(* IEC 61131-3 sources: llm-plc-st-eval/codesys/dobles/B2, 5 files *)

(* ---- 01_Correcta.st ---- *)
(* DOBLE DE PRUEBA B2/Correcta - NO ES CORPUS. Esperado: veredicto 1 *)
FUNCTION_BLOCK FB_Valvula
VAR_INPUT
    nivelAlto : BOOL;
END_VAR
VAR_OUTPUT
    valvula : BOOL;
END_VAR
VAR
    t : TON;
END_VAR
t(IN := nivelAlto, PT := T#5S);
valvula := t.Q;
END_FUNCTION_BLOCK

(* ---- 02_TofEnVezDeTon.st ---- *)
(* DOBLE DE PRUEBA B2/TofEnVezDeTon - NO ES CORPUS. Esperado: veredicto 2, falla en el paso 1 *)
FUNCTION_BLOCK FB_Valvula
VAR_INPUT
    nivelAlto : BOOL;
END_VAR
VAR_OUTPUT
    valvula : BOOL;
END_VAR
VAR
    t : TOF;
END_VAR
t(IN := nivelAlto, PT := T#5S);
valvula := t.Q;
END_FUNCTION_BLOCK

(* ---- 03_PresetCorto.st ---- *)
(* DOBLE DE PRUEBA B2/PresetCorto - NO ES CORPUS. Esperado: veredicto 2, falla en el paso 1 *)
FUNCTION_BLOCK FB_Valvula
VAR_INPUT
    nivelAlto : BOOL;
END_VAR
VAR_OUTPUT
    valvula : BOOL;
END_VAR
VAR
    t : TON;
END_VAR
t(IN := nivelAlto, PT := T#2S);
valvula := t.Q;
END_FUNCTION_BLOCK

(* ---- 04_SinCierreInmediato.st ---- *)
(* DOBLE DE PRUEBA B2/SinCierreInmediato - NO ES CORPUS. Esperado: veredicto 2, falla en el paso 3 *)
FUNCTION_BLOCK FB_Valvula
VAR_INPUT
    nivelAlto : BOOL;
END_VAR
VAR_OUTPUT
    valvula : BOOL;
END_VAR
VAR
    t : TON;
END_VAR
t(IN := nivelAlto, PT := T#5S);
IF t.Q THEN
    valvula := TRUE;
END_IF
END_FUNCTION_BLOCK

(* ---- 05_UnSoloDisparo.st ---- *)
(* DOBLE DE PRUEBA B2/UnSoloDisparo - NO ES CORPUS. Esperado: veredicto 2, falla en el paso 4 *)
FUNCTION_BLOCK FB_Valvula
VAR_INPUT
    nivelAlto : BOOL;
END_VAR
VAR_OUTPUT
    valvula : BOOL;
END_VAR
VAR
    t : TON;
    yaAbrio : BOOL;
END_VAR
t(IN := nivelAlto, PT := T#5S);
IF t.Q AND NOT yaAbrio THEN
    valvula := TRUE;
    yaAbrio := TRUE;
END_IF
IF NOT nivelAlto THEN
    valvula := FALSE;
END_IF
END_FUNCTION_BLOCK
